(* IEC 61131-3 sources: Jacob-Formschaumtechnik-ISEL-CNC-Retrofit/twincat/PLC/src/2_Devices, 2 files *)

(* ---- FB_AxisSupervisor.st ---- *)
(* Ueberwacht vier Achsen (Index 1..4) und fasst Zustaende fuer die Meldeliste zusammen.
   Muss-Anforderungen: 2.2.3 Hardware-Endschalter, 2.2.6 Referenzverlust, 2.10.4 Ueberwachung
   von Feldbus und Antrieben. Endschalter im Ruhestrom (FALSE = ausgeloest). *)
FUNCTION_BLOCK FB_AxisSupervisor
VAR_INPUT
    bEnableCmd      : BOOL;     (* Reglerfreigabe angefordert *)
    bFieldbusOk     : BOOL;
    bHomingActive   : BOOL;     (* gewollte Referenzfahrt laeuft: kein Referenzverlust (Befund 5) *)
    rMaxFollowErr   : LREAL;    (* mm, [Annahme] bis Achsdaten vorliegen *)
END_VAR
VAR_IN_OUT
    aAxis : ARRAY[1..4] OF ST_AxisDrive;
END_VAR
VAR_OUTPUT
    bAnyFault      : BOOL;
    bAnyHwLimit    : BOOL;
    bFollowErr     : BOOL;
    bAllReady      : BOOL;
    bAllEnabled    : BOOL;
    bAllHomed      : BOOL;
    bHomingLost    : BOOL;      (* Referenz war da und ist weg (Regler aus/Fehler) *)
    bEnableTimeout : BOOL;      (* Freigabe angefordert, aber Antriebe melden nicht freigegeben (Befund 14) *)
END_VAR
VAR
    i           : INT;
    bHadHomed   : BOOL;
    tonEnable   : TON;
END_VAR

bAnyFault := FALSE; bAnyHwLimit := FALSE; bFollowErr := FALSE;
bAllReady := TRUE; bAllEnabled := TRUE; bAllHomed := TRUE;

FOR i := 1 TO 4 DO
    IF aAxis[i].bFault THEN bAnyFault := TRUE; END_IF
    IF NOT aAxis[i].bHwLimitPlus OR NOT aAxis[i].bHwLimitMinus THEN bAnyHwLimit := TRUE; END_IF
    IF ABS(aAxis[i].rFollowErr) > rMaxFollowErr THEN bFollowErr := TRUE; END_IF
    IF NOT aAxis[i].bReady   THEN bAllReady := FALSE; END_IF
    IF NOT aAxis[i].bEnabled THEN bAllEnabled := FALSE; END_IF
    IF NOT aAxis[i].bHomed   THEN bAllHomed := FALSE; END_IF
END_FOR

(* Referenzverlust: war referenziert und ist es nicht mehr *)
IF bAllHomed THEN
    bHadHomed := TRUE;
    bHomingLost := FALSE;
ELSIF bHomingActive THEN
    bHadHomed := FALSE;
    bHomingLost := FALSE;
ELSIF bHadHomed THEN
    bHomingLost := TRUE;
    bHadHomed := FALSE;
END_IF
IF NOT bFieldbusOk THEN
    bAllReady := FALSE; bAllEnabled := FALSE;
END_IF

tonEnable(IN := bEnableCmd AND bFieldbusOk AND NOT bAllEnabled, PT := T#3S);
bEnableTimeout := tonEnable.Q;
END_FUNCTION_BLOCK

(* ---- FB_Spindle.st ---- *)
(* Spindel isel VKH63/26-90T, 2,2 kW, max. 16600 1/min, am FU Emerson Commander SK.
   Ansteuerung Variante 1: Start/Richtung digital, Drehzahl 0..10 V. Variante Modbus RTU ist offen.
   [Annahme] Start und Richtung als getrennte Ausgaenge, FU-Rueckmeldung "bereit" und "Drehzahl erreicht"
   als Eingaenge. Bis Schaltplan vorliegt, ist das nicht belegt.
   Befund 1 der Papierpruefung: Die Anforderung ist selbsthaltend. Ein Start entsteht nur aus einer
   steigenden Flanke von bStartCw/bStartCcw. Jeder Stopp (Release weg, Fehler, bStop, Einrichten)
   loescht die Anforderung. Ein noch anstehender Pegel startet die Spindel nie von selbst neu.
   Befund 13: Drehrichtungsumkehr nur ueber Stillstand (Auslaufzeit). *)
FUNCTION_BLOCK FB_Spindle
VAR_INPUT
    bRelease      : BOOL;        (* Betriebsart + Sicherheit erlauben die Spindel *)
    bSetupLocked  : BOOL;        (* Betriebsart Einrichten/Test: Spindel gesperrt *)
    bStop         : BOOL;        (* Stopp-Anforderung (Abbruch, R3/R4, NOT-HALT): loescht die Anforderung *)
    bStartCw      : BOOL;        (* M3 bzw. Hand-Taste, Pegel *)
    bStartCcw     : BOOL;        (* M4 bzw. Hand-Taste, Pegel *)
    rSetRpm       : REAL;        (* S-Wert, 1/min *)
    rOverridePct  : REAL;        (* 0..150 *)
    bFuReady      : BOOL;        (* FU bereit, Ruhestrom: FALSE = Stoerung *)
    bFuAtSpeed    : BOOL;        (* [Annahme] FU meldet Drehzahl erreicht *)
    bPtcOk        : BOOL;        (* Kaltleiter Motor, Ruhestrom: FALSE = Uebertemperatur *)
    bAckReset     : BOOL;
    rMaxRpm       : REAL;
    rMinRpm       : REAL;
    rVoltMax      : REAL;
    tRunUp        : TIME;
    tStandstill   : TIME;
    bAllowPend    : BOOL := TRUE; (* G-11: Start darf auf Stillstand warten (Programm). FALSE (Hand): Start waehrend des Auslaufs wird verworfen *)
END_VAR
VAR_OUTPUT
    bRunCmd       : BOOL;        (* Ausgang Start *)
    bDirCcw       : BOOL;        (* Ausgang Richtung *)
    rVoltOut      : REAL;        (* Ausgang 0..10 V (EL4002) *)
    bRunning      : BOOL;        (* Drehzahl erreicht *)
    bStandstillOk : BOOL;        (* Spindel steht (Auslaufzeit abgelaufen) *)
    bFault        : BOOL;
    bPtcTrip      : BOOL;
    bNoFeedback   : BOOL;
    bLockedSetup  : BOOL;        (* Start versucht, aber gesperrt *)
    rActRpm       : REAL;        (* berechneter Sollwert nach Override; kein Istwert! *)
END_VAR
VAR
    tonRunUp   : TON;
    tonStop    : TON;
    rRpm       : REAL;
    bWantRun   : BOOL;
    bLatchFault: BOOL;
    rtAck      : R_TRIG;
    rtCw       : R_TRIG;
    rtCcw      : R_TRIG;
    nDirAct    : INT;            (* 0 = keine Anforderung, 1 = rechts, 2 = links *)
    nDirPend   : INT;            (* wartet auf Stillstand, 0 = nichts *)
    bStopCond  : BOOL;
    bSpeedInvalid : BOOL;        (* G-12: Start ohne gueltigen S-Wert *)
END_VAR

rtAck(CLK := bAckReset);
rtCw(CLK := bStartCw);
rtCcw(CLK := bStartCcw);

bPtcTrip := NOT bPtcOk;
bFault   := NOT bFuReady OR bPtcTrip;
IF bFault THEN bLatchFault := TRUE; END_IF
IF bLatchFault AND rtAck.Q AND bFuReady AND bPtcOk THEN bLatchFault := FALSE; END_IF

bLockedSetup := bSetupLocked AND (bStartCw OR bStartCcw);

(* Anforderung verwalten *)
bStopCond := bStop OR NOT bRelease OR bSetupLocked OR bLatchFault;
IF bStopCond THEN
    nDirAct := 0; nDirPend := 0;
ELSE
    (* Ende der Anforderung: M5 bzw. Taste aus *)
    IF NOT bStartCw  AND nDirAct = 1 THEN nDirAct := 0; END_IF
    IF NOT bStartCcw AND nDirAct = 2 THEN nDirAct := 0; END_IF
    IF NOT bStartCw  AND nDirPend = 1 THEN nDirPend := 0; END_IF
    IF NOT bStartCcw AND nDirPend = 2 THEN nDirPend := 0; END_IF
    (* neuer Start nur mit steigender Flanke *)
    IF rtCw.Q  AND bStartCw  AND NOT bStartCcw AND (bAllowPend OR bStandstillOk) THEN nDirPend := 1; END_IF
    IF rtCcw.Q AND bStartCcw AND NOT bStartCw  AND (bAllowPend OR bStandstillOk) THEN nDirPend := 2; END_IF
    (* Start erst, wenn die Spindel steht (auch bei Richtungsumkehr) *)
    IF nDirPend <> 0 AND nDirAct = 0 AND bStandstillOk THEN
        nDirAct := nDirPend; nDirPend := 0;
    END_IF
END_IF

bWantRun := nDirAct <> 0;
(* G-12: Kein gueltiger S-Wert (0 oder fehlt): Spindel nicht anfahren, Meldung 202 (R3) *)
bSpeedInvalid := bWantRun AND rSetRpm <= 0.0;
bRunCmd  := bWantRun AND NOT bSpeedInvalid;
bDirCcw  := nDirAct = 2;

(* Drehzahl begrenzen und Override anwenden *)
rRpm := rSetRpm * LIMIT(0.0, rOverridePct, 150.0) / 100.0;
rRpm := LIMIT(rMinRpm, rRpm, rMaxRpm);
IF bRunCmd AND rMaxRpm > 0.0 THEN
    rVoltOut := rRpm / rMaxRpm * rVoltMax;
    rActRpm  := rRpm;
ELSE
    rVoltOut := 0.0;
    rActRpm  := 0.0;
END_IF

(* Rueckmeldung: nach Hochlaufzeit muss FU "Drehzahl erreicht" melden *)
tonRunUp(IN := bWantRun, PT := tRunUp);
bRunning    := bWantRun AND bFuAtSpeed;
bNoFeedback := (tonRunUp.Q AND NOT bFuAtSpeed) OR bSpeedInvalid;

(* Auslaufzeit: Stillstand gilt erst nach Ablauf *)
tonStop(IN := NOT bWantRun, PT := tStandstill);
bStandstillOk := tonStop.Q;
END_FUNCTION_BLOCK
